// TIA Portal V20 export
FUNCTION "Störmeldungen" : Void   // FC512, STL
TITLE = Störmeldungen
{ S7_Optimized_Access := 'FALSE' }
// Störmeldungsbaustein: Hier befinden sich alle Störungen zusammengefasst zur 
// Sammelstörung und alle Störungen, die nicht in FB`s aufgelistet wurden.
// stored: AutoNumber false
   VAR_TEMP
      retval : Int;
      keine_Störung : Bool;
   END_VAR
BEGIN

NETWORK
TITLE = Sammelstörung Anlage
      A     "ProDiag_Allgemein_DB".State.C1;
      O     "POS3_0_Prodiag_DB".State.C1;



// Schrittketten in Störung (Interlock oder Supervision)
      O     "POS3_0_Signal".Schrittkette.ERR_FLT;

      =     "HMI_Signale".Sammelstoerung;


NETWORK
TITLE = Stop von Störmeldungen



      CLR;
      S     "HMI_Signale".Stop_Von_Stoermeldung;

      A     "03_Betriebsart_DB".ACK_Taste;
      R     "HMI_Signale".Stop_Von_Stoermeldung;
END_FUNCTION
